(* IEC 61131-3 sources: Elmo_Master/Lasal_PRG/Welcon8Axis_EtherCAT_Test_With_RobotAxis/Network/Robot_Network, 1 file *)

(* ---- ONE_Robot_Network_Table.st ---- *)
#define OBJECTS_CONFIG

//Define part of class _LMCBeltAxis
//#define _DEBUG_MODUS_ISSYNCHRON
//#define _DEBUG_MODUS_CHECKSWLIMIT

#define _LMCBELT_MIN_POS       -16#6FFFFFFF    // default MINPOS when INITvalue=0
#define _LMCBELT_MAX_POS        16#6FFFFFFF    // default MAXPOS when INITvalue=0
#define _LMCBELT_OVERVFLOW_POS  16#7FFFFFFF    // MAX POSITION for checking overflow

#define _LMCBELT_AMAX_SET 2000000000
#define _LMCBELT_VMAX_SET 500000000

//////////////////////
// ruckbegrenzter Modus _JERK_PROFILE
#define LMCBELT_MIN_SHRINK_FACTOR_4_CORRECTTOEXACTPOS 0.9
#define LMCBELT_MAX_SHRINK_FACTOR_4_CORRECTTOEXACTPOS_FAR 1.2
#define LMCBELT_MAX_SHRINK_FACTOR_4_CORRECTTOEXACTPOS_NEAR 5.0
#define LMCBELT_MAX_SHRINK_FACTOR_4_CORRECTTOEXACTPOS_WINDOW 5.0

#define LMCBELT_MAX_TIME_TO_WAIT_4_BRAKING 3.0 //in Ticks
#define LMCBELT_MAX_DURATION_WITH_MAX_ACCEL_TO_MASTER 20000  //in Ticks
#define LMCBELT_ALLOWED_AJMP_FACTOR 1.1
#define LMCBELT_FACTOR_4_ALLOWED_MASTER_ACCEL_PROFILE_COUPLING 1.2
#define LMCBELT_ACCEL_FACTOR_4_PROFILE_COUPLING 1.1
#define LMCBELT_JERK_FACTOR_4_PROFILE_COUPLING 1.2
#define LMCBELT_FACTOR_2_REDUCE_AXIS_ACC_LIMIT 1.02

//////////////////////
// LREAL Modi
// #define DEBUG_TRAP_DELTA_ACCEL
#define _LMCBELT_LREAL_EPSILON 0.000001

#ifndef _DINT_MIN
#define _DINT_MIN -2147483648
#endif

#ifndef _DINT_MAX
#define _DINT_MAX 2147483647
#endif

#define _LMCBELT_MIN_VEL_MOVECMD 1 // minimale programmierbare Geschwindigkeit für LREAL-MoveTypes [internal units / sec]
#include <.\lsl_st_systrace.h>
#include "..\..\Class\_LMCAxisBase\C_MathAxis.h"
#include "..\..\Class\_LMCAxisBase\_LMCTraceView.h"
//Define part of class _LMCMath_SO3
// maximal inaccuracies of LREAL
#define _LREAL_EPSILON        0.000001
#define _LREAL_EPSILON_MUL    0.000001
// minmal volume of orthogonalsystem
#define MIN_SPAT_PRODUCT      _LREAL_EPSILON_MUL

#ifndef deg
  #define SCALE_ROT_ANGLE       (10000)
#else
  #define SCALE_ROT_ANGLE       (1deg)
#endif

#define SCALE_VECTOR          (10000)
//Define part of class _LMCMathFunctions
#define _INT_DEG                       * 1024 * 1000 //Internal Resolution of Degrees
#define LMC_PI                          3.1415926535897932384626433832795   //LMC_ avoids name clash

#define _LMC_EPSILON    0.000001
#define _MATH_EPSILON   0.000000001

//LREAL Zero Test:
#ifndef _LMCMATH_FLOAT_ISZERO
  #define _LMCMATH_FLOAT_ISZERO(p1)            ((p1 > -_LMC_EPSILON) & (p1 < _LMC_EPSILON))
#endif
#ifndef _LMCMATH_FLOAT_NOTZERO
  #define _LMCMATH_FLOAT_NOTZERO(p1)           ((p1 < -_LMC_EPSILON) | (p1 > _LMC_EPSILON))
#endif
#ifndef _LMCMATH_FLOAT_EQUAL
  #define _LMCMATH_FLOAT_EQUAL(p1,p2)          (((p1 - p2) < _LMC_EPSILON) & ((p1 - p2) > -_LMC_EPSILON))
#endif

#define _LMCMATH_LREAL_MAX  1.79E308
#define _LMCMATH_REAL_MAX   3.4E38

#ifndef _DINT_MIN
  #define _DINT_MIN -2147483648
#endif

#define LMC_NUMERIC_TOLERANCE   (0.000000001)
#define LMC_RESOLVE_TOLERANCE       (0.000000001)

// 25µsec für ein repeat auf ARM CP 111
#define LMC_MAX_REPEAT      25

// Geschwindigkeit wird auf 1 interne Einheit genau iteriert
#define PRECIS_REPEAT   (1.0)

//#define INTERN_MATH_TEST
#include "..\..\Class\_LMCMathFunctions\C_MathFunct.h"
//Define part of class _LMCProfileBase
#pragma once

// DEBUG MODUS TO DEACTIVATE ACTIVE MUTEX
//#define DEBUG_MODUS
//#define DEBUG_CMD_TYPE

#pragma once

//LREAL Zero Test:
#ifndef _LMCPROF_LREAL_ISZERO
  #define _LMCPROF_LREAL_ISZERO(p1)           ((p1 > -_LMCPROF_EPSILON) & (p1 < _LMCPROF_EPSILON))
#endif
#ifndef _LMCPROF_LREAL_NOTZERO
  #define _LMCPROF_LREAL_NOTZERO(p1)          ((p1 < -_LMCPROF_EPSILON) | (p1 > _LMCPROF_EPSILON))
#endif
#define _LMCPROF_LREAL_MAX                    1.79E308

#define _LMPROF_PROMILLE                      1000

//Move Curve Spline Defines
#define _LMC_PROF_MCS_MINOVERDRIVE                -900
#define _LMC_PROF_MCS_MAXOVERDRIVE                10000 //=> Centripetal Acceleration can be up to 10 * given AMove
#define _LMC_PROF_MCS_DEFAULT_JERKSMOOTH          1

#define _LMC_PROF_CES_DEFAULT_ZEXPONENT           1.0 //Default Spline Z Exponent used in calcEllipseSpline(), set with SetProfileParameter()
#define _LMC_PROF_CES_MAX_ZEXPONENT_W_LIN         1.0 //Max Spline Z Exponent if moving with Linear movements, used in calcEllipseSpline()
#define _LMC_PROF_CES_MIN_ZEXPONENT               1.0 //Min Spline Z Exponent, used in calcEllipseSpline()

#define _LMC_PROF_ERRORBUFFER_ENTRIES             10
#define _LMC_PROF_MAINGROUP                       1 // Achse ist in Hauptgruppe
#define _LMC_PROF_SLAVEGROUP1                     2 // Achse ist in Nebengruppe 1
#define _LMC_PROF_SLAVEGROUP2                     3 // Achse ist in Nebengruppe 2
#define _LMC_PROF_SLAVEGROUP3                     4 // Achse ist in Nebengruppe 3
#define _LMC_PROF_SLAVEGROUP4                     5 // Achse ist in Nebengruppe 4
#define _LMC_PROF_SLAVEGROUP5                     6 // Achse ist in Nebengruppe 5

#define _LMC_PROF_MAX_SLAVEGROUPS               _LMC_PROF_SLAVEGROUP5

#define _LMCPROF_NEEDED_FREE_BUFFER_ENTRIES    4

#define _LMC_PROF_MAXOVERRIDE	               1000 // Maximalwert für Override
#define _LMC_PROF_MINOVERRIDE	                  0	// Minimalwert für Override
#define _LMC_PROF_NORMOVERRIDE               1000 // 100%-Wert für Override

#define _LMC_PROF_MAX_DINT                   2147483647
#define _LMC_PROF_MAX_UDINT                  4294967295

#define TRANS1                                  0 //index of 1. transition elmt
#define TRANS2                                  1 //index of 2. transition elmt
#define TRANS3                                  2 //index of 3. transition elmt

#define _LMC_PROF_VECTOR_WINDOW                 10mm

#define MIN_TRANSRAD_PPTH                       0
#define DEF_TRANSRAD_PPTH                       500
#define MOVECURVE_ACCEL_PATH_AUXAXIS            250 // 250 // 25% of the path length is used for accelerating auxiliary axes with splines

#define _LMC_PROF_DEFAULT_MAX_TANG_ERR          900000 //90° ist defaultmäßig maximale tangential fehler

#define _LMC_PROF_RESTARTPROF_TOLSPHERE_DEFAULT 1mm
#define _LMC_PROF_RESTARTPROF_APPROACH_DEFAULT  0

#define _LMC_PROF_MULT_LOOKAHEAD_LINE           5 //default multiplier for lookaheadsmalllines

#define _LMCPROF_REDUCEMOVINGTIME_MAXFACTOR  10000

// the minimal height difference between the end / beginning of the linear part of a MoveCurve() movement and the start / end of the MoveCurveAux section
#define _LMCPROF_MINIMAL_SWERVEDIFF            0.2mm

// Fehlertoleranz bei Umrechnung von Integer auf Float
#define RESOLUTION_ERROR      (5.0)
// Fehlertoleranz wenn der Ruck innerhalb eines Ticks um 2*Jmax springt
#define JERKTICK_ERROR        (-1.0)

// Rückgabeparameter
#define CALCRESIDT_NO_ERROR            0
#define CALCRESIDT_INIT_ERROR          -1
#define CALCRESIDT_NO_SOLUTION         -2

// Präfix (wird für Ruck verwendet)
#ifndef PREFIX_KILO
  #define PREFIX_KILO             (1000.0)
#endif
// Umrechnung von Sekunden auf Ticks
#ifndef CONVERT_SEC_TO_MSEC
  #define CONVERT_SEC_TO_MSEC   (1000.0)
#endif
// interne Mathematik-Tests - speziell Genauigkeitstest von LREAL
//#define INTERN_TEST

// =======================================================
// Defines for Clothoid (Parameters / Conversion)
// Minimal angle to use a compound solution
#define _LMCPROF_CLOTH_MINTAU                  0.06        // 0.06 (radiant) = R/3 clothoid identification
#define _LMCPROF_CLOTH_HAIRPINLIMIT            0.0004      // 0.0004 (radiant) < 0.025 degree - Limit, when the turn is close to a hairpin (cone angle smaller than this limit - handle it is a stop)
#define _LMCPROF_CLOTH_TABLESCALE              0.000000001 // 10^(-9) // This value is a fixed scale of the unit cloth table - when this value is changed, the table must be changed too.

//Angle conversion
#ifndef _LMCPROF_DEG_RAD
  #define _LMCPROF_DEG_RAD(p1)       (((p1) / (180.0 * 1deg)) * _PI)
#endif
#ifndef _LMCPROF_RAD_DEG
  #define _LMCPROF_RAD_DEG(p1)       (((p1) / _PI) * 180.0) * 1deg
#endif

// Defines for tangential axis
#define _LMCPROF_TANGAXIS_ACTANGLEOVERFLOWLIMIT    45.0 deg
#define _LMCPROF_TANGAXIS_OVERFLOWDETECTLIMIT     359.0 deg

// Maximum allowed number of points per spline -
// Attention! If this value is changed also the MaxNrOfPointsPerMoveMaxValue of MoveSplineTable and
// IPR_MAX_NR_SPLINE_POINTS of _LMCCNCIPRBase are to be changed
#define PROF_MAX_NR_SPLINE_POINTS           50
// Maximal number of spline points is twice as high as the number of points - 1 (movement to the last point can't include addition intermediate move)
#define PROF_MaxNrSplineTargets             ((PROF_MAX_NR_SPLINE_POINTS * 2) - 1)

// Move Spline minimal trajectory angle
#define _LMC_PROF_MOVESPLINE_MIN_ANGLE      45 deg // 45 deg
#include "..\..\Class\_LMCProfileBase\C_MathProfile.h"
//Define part of class _LMCProfileBuffer
#define    _LMC_PB_MINENTRIES     201
#define    _LMC_PB_MAXENTRIES     2000

#define _LMC_PB_TMP_MINENTRIES    7
#define _LMC_PB_TMP_MAXENTRIES    100

#define _LMC_PB_RB_MINENTRIES     5
#define _LMC_PB_RB_MAXENTRIES     10

//////////////////////
// Mutex
#define MUTEX_NAME_MAX_LENGTH_LMCPROFILE     32   //maximale Anzahl an Zeichen für den Mutexnamen
#define MUTEX_NAME_END_LENGTH_LMCPROFILE      3
#define STR_MUTEX_NAME_SEPERATOR_LMCPROFILE ".."
//Define part of class _LMCRobotBase
#define DELAYPOWERONHWAXES_TIMEOUT        0
#define DELAYPOWEROFF_TIMEOUT             0
#define WAITPOWERONHWAXES_TIMEOUT     30sec
#define CHECKREFERENCEHWAXES_TIMEOUT  30sec
#define WAITPOWERONKINAXES_TIMEOUT    30sec
#define CHECKCOUPLEHWAXES_TIMEOUT        50
#define WAITPROFILESTOPPED_TIMEOUT     1000
#define WAITSTOPMOVEKINAXES_TIMEOUT    1000
#define WAITSTOPMOVEHWAXES_TIMEOUT     1000
#define WAITERRORQUIT_TIMEOUT           800

#define STOPMOVEPOSITIONWINDOW_DEFAULT 1mm
#define START_COUPLEWINDOW_DEFAULT     1mm

#define GET_LINE_OFFSET 1000000

#define ALL_HW_AXES -1
#define ALL_KINEMATIC_AXES -2
#define ALL_PROFILE_AXES -3
#define ALL_AXES_101_TO_109 -4
#define ALL_ROBOT_AXES 0

#define SCALE_ROTAXIS 100000
#define SCALE_KOFAC 1000000

#define LIMIT_BELT_CMD            2
#define SYNC_DESYNC_FULL_LENGTH   1000

#define SYNC_DESYNC_MIN_LENGTH      50

#define BELTCOUPLING_DEFAULT_FILTER_DEPTH_VMASTER 40 //Bei Änderungen auch Kommentar von _LMCROBOT_BELTCOUPLING_VEL_FILTER_DEPTH anpassen!
#define BELTCOUPLING_MAX_FILTER_DEPTH_VMASTER 60 //Bei Änderungen auch Kommentar von _LMCROBOT_BELTCOUPLING_VEL_FILTER_DEPTH anpassen!

#define ROTATORY_DISK_MODULO (360deg)
#define ROTATORY_DISK_ANGLE_TO_RADIANT (2.0*LMC_PI/(ROTATORY_DISK_MODULO))

#ifndef CIRCLE3D_NO_HELIX_MAX_DEVIATION
  #define CIRCLE3D_NO_HELIX_MAX_DEVIATION 0.02
#endif
//Define part of class _LMCSplineBuffer
#define LMCSPLINEBUFF_MINBUFFS              3             //SplineGroups
#define LMCSPLINEBUFF_EPSILON               0.000001
#define LMCSPLINEBUFF_MAX_SPLINES_PER_GROUP 40
#define LMCSPLINEBUFF_MALLOC_MARK           9
#define LMCSPLINEBUFF_HIRES_VEL_DEFAULT     (1000.0)
#define LMCSPLINEBUFF_HIRES_ACC_DEFAULT     (10000.0)
#define LMCSPLINEBUFF_HIRES_JERK_DEFAULT    (1000000.0)
#define LMCSPLINEBUFF_CALCPARAS_POS         16#00000001
#define LMCSPLINEBUFF_CALCPARAS_VEL         16#00000002
#define LMCSPLINEBUFF_CALCPARAS_ACC         16#00000004
#define LMCSPLINEBUFF_CALCPARAS_JERK        16#00000008
#define LMCSPLINEBUFF_CALCPARAS_JOUNCE      16#00000010
#define LMCSPLINEBUFF_SEARCH_ITER_DEFAULT   100
#define LMCSPLINEBUFF_SEARCH_WIN_DEFAULT    1.0

//Coeffecient Short Names:
#define SB_CO_A (pSplineSection^.Coefficients.lrCoefficient1)
#define SB_CO_B (pSplineSection^.Coefficients.lrCoefficient2)
#define SB_CO_C (pSplineSection^.Coefficients.lrCoefficient3)
#define SB_CO_D (pSplineSection^.Coefficients.lrCoefficient4)
#define SB_CO_E (pSplineSection^.Coefficients.lrCoefficient5)
#define SB_CO_F (pSplineSection^.Coefficients.lrCoefficient6)
#define SB_CO_G (pSplineSection^.Coefficients.lrCoefficient7)
#define SB_CO_H (pSplineSection^.Coefficients.lrCoefficient8)
#define SB_TICK (pSplineSection^.lrTick)
//Define part of class _LMCTableBuffer
#define _TABLE_POINT_COUNT_ 100

#define _TABLE_POINT_20PERCENT 25
#define _TABLE_POINT_35PERCENT 40
#define _TABLE_POINT_50PERCENT 50
#define _TABLE_POINT_65PERCENT 60
#define _TABLE_POINT_80PERCENT 75

#define _LMCTABLEBUFFER_MALLOCMARK  9

FUNCTION GLOBAL TAB ONE_Robot_Network
-1$UINT, 0$UINT,
0$UINT, 0$UINT,

16$UDINT,
TO_UDINT(1064285160), "_LMCBeltAxis", 1$UINT, 7$UINT, 1$UINT,
TO_UDINT(4293818033), "_LMCMath_SO3", 1$UINT, 24$UINT, 2$UINT,
TO_UDINT(838927485), "_LMCMathFunctions", 1$UINT, 75$UINT, 2$UINT,
TO_UDINT(2952189205), "_LMCProfile", 3$UINT, 0$UINT, 0$UINT,
TO_UDINT(506182625), "_LMCProfileBase", 4$UINT, 0$UINT, 0$UINT,
TO_UDINT(2726627155), "_LMCProfileBuffer", 1$UINT, 53$UINT, 1$UINT,
TO_UDINT(2883857672), "_LMCProfileLog", 1$UINT, 44$UINT, 1$UINT,
TO_UDINT(4141185109), "_LMCProfileVis", 1$UINT, 30$UINT, 1$UINT,
TO_UDINT(3174746949), "_LMCProfileVisAxis", 1$UINT, 20$UINT, 9$UINT,
TO_UDINT(4192117043), "_LMCProfileVisInt", 1$UINT, 41$UINT, 1$UINT,
TO_UDINT(1543035932), "_LMCProfileVisMovePara", 1$UINT, 30$UINT, 6$UINT,
TO_UDINT(3888346726), "_LMCRobotBase", 2$UINT, 22$UINT, 1$UINT,
TO_UDINT(4210476436), "_LMCRobotLog", 1$UINT, 42$UINT, 1$UINT,
TO_UDINT(1286231841), "_LMCSplineBuffer", 1$UINT, 2$UINT, 1$UINT,
TO_UDINT(2328372307), "_LMCTableBuffer", 1$UINT, 23$UINT, 1$UINT,
TO_UDINT(1472648579), "Robot_Handler", 0$UINT, 0$UINT, 1$UINT,

1$UINT, TO_UDINT(3188917884), "_LMCROBOTBASE1\LMCBELTINTERNAL",

1$UINT, TO_UDINT(2922016232), "_LMCROBOTBASE1\LMCMATH_SO3",
1$UINT, TO_UDINT(1366148008), "_LMCROBOTBASE1\_BASE\_LMCMATH_SO3",

1$UINT, TO_UDINT(1157192838), "_LMCROBOTBASE1\LMCBELTINTERNAL\LMCMATH",
1$UINT, TO_UDINT(2796190616), "_LMCROBOTBASE1\_BASE\_LMCMATHFUNCTIONS",

1$UINT, TO_UDINT(909015222), "_LMCROBOTBASE1\_BASE\_LMCPROFILEBUFFER",

1$UINT, TO_UDINT(2347724176), "_LMCROBOTBASE1\_BASE\_LMCPROFILELOG",

1$UINT, TO_UDINT(3604887757), "_LMCROBOTBASE1\_BASE\_LMCPROFILEVIS",

1$UINT, TO_UDINT(4143639116), "_LMCROBOTBASE1\_BASE\_LMCPROFILEVIS\_LMCPROFILEVISAXIS1",
1$UINT, TO_UDINT(1878244342), "_LMCROBOTBASE1\_BASE\_LMCPROFILEVIS\_LMCPROFILEVISAXIS2",
1$UINT, TO_UDINT(418679648), "_LMCROBOTBASE1\_BASE\_LMCPROFILEVIS\_LMCPROFILEVISAXIS3",
1$UINT, TO_UDINT(2257592003), "_LMCROBOTBASE1\_BASE\_LMCPROFILEVIS\_LMCPROFILEVISAXIS4",
1$UINT, TO_UDINT(4053216853), "_LMCROBOTBASE1\_BASE\_LMCPROFILEVIS\_LMCPROFILEVISAXIS5",
1$UINT, TO_UDINT(1755217903), "_LMCROBOTBASE1\_BASE\_LMCPROFILEVIS\_LMCPROFILEVISAXIS6",
1$UINT, TO_UDINT(530141049), "_LMCROBOTBASE1\_BASE\_LMCPROFILEVIS\_LMCPROFILEVISAXIS7",
1$UINT, TO_UDINT(2401653480), "_LMCROBOTBASE1\_BASE\_LMCPROFILEVIS\_LMCPROFILEVISAXIS8",
1$UINT, TO_UDINT(4162937470), "_LMCROBOTBASE1\_BASE\_LMCPROFILEVIS\_LMCPROFILEVISAXIS9",

1$UINT, TO_UDINT(2979030242), "_LMCROBOTBASE1\_BASE\_LMCPROFILEVIS\_LMCPROFILEVISINT",

1$UINT, TO_UDINT(1783828595), "_LMCROBOTBASE1\_BASE\_LMCPROFILEVIS\_LMCPROFILEVISMOVEPARA1",
1$UINT, TO_UDINT(4082778569), "_LMCROBOTBASE1\_BASE\_LMCPROFILEVIS\_LMCPROFILEVISMOVEPARA2",
1$UINT, TO_UDINT(2220716383), "_LMCROBOTBASE1\_BASE\_LMCPROFILEVIS\_LMCPROFILEVISMOVEPARA3",
1$UINT, TO_UDINT(440001788), "_LMCROBOTBASE1\_BASE\_LMCPROFILEVIS\_LMCPROFILEVISMOVEPARA4",
1$UINT, TO_UDINT(1832834154), "_LMCROBOTBASE1\_BASE\_LMCPROFILEVIS\_LMCPROFILEVISMOVEPARA5",
1$UINT, TO_UDINT(4097279440), "_LMCROBOTBASE1\_BASE\_LMCPROFILEVIS\_LMCPROFILEVISMOVEPARA6",

_NO_ATTR, TO_UDINT(669706412), "_LMCROBOTBASE1",

1$UINT, TO_UDINT(2991295094), "_LMCROBOTBASE1\_LMCROBOTLOG",

1$UINT, TO_UDINT(2213426856), "_LMCROBOTBASE1\_BASE\_LMCSPLINEBUFFER",

1$UINT, TO_UDINT(1950102629), "_LMCROBOTBASE1\_BASE\_LMCTABLEBUFFER",

_NO_ATTR, TO_UDINT(4147837944), "ROBOT_HANDLER1",

//Internal connections
0$UDINT,
27$UDINT,
TO_UDINT(0), "LMCMath", TO_UDINT(3),
TO_UDINT(7), "_LMCProfileVisMovePara1", TO_UDINT(18),
TO_UDINT(7), "_LMCProfileVisMovePara2", TO_UDINT(19),
TO_UDINT(7), "_LMCProfileVisMovePara3", TO_UDINT(20),
TO_UDINT(7), "_LMCProfileVisMovePara4", TO_UDINT(21),
TO_UDINT(7), "_LMCProfileVisMovePara5", TO_UDINT(22),
TO_UDINT(7), "_LMCProfileVisMovePara6", TO_UDINT(23),
TO_UDINT(7), "_LMCProfileVisAxis1", TO_UDINT(8),
TO_UDINT(7), "_LMCProfileVisAxis2", TO_UDINT(9),
TO_UDINT(7), "_LMCProfileVisAxis3", TO_UDINT(10),
TO_UDINT(7), "_LMCProfileVisAxis4", TO_UDINT(11),
TO_UDINT(7), "_LMCProfileVisAxis5", TO_UDINT(12),
TO_UDINT(7), "_LMCProfileVisAxis6", TO_UDINT(13),
TO_UDINT(7), "_LMCProfileVisInt", TO_UDINT(17),
TO_UDINT(7), "_LMCProfileVisAxis7", TO_UDINT(14),
TO_UDINT(7), "_LMCProfileVisAxis8", TO_UDINT(15),
TO_UDINT(7), "_LMCProfileVisAxis9", TO_UDINT(16),
TO_UDINT(24), "_LMCMathFunctions", TO_UDINT(4),
TO_UDINT(24), "_LMCProfileBuffer", TO_UDINT(5),
TO_UDINT(24), "_LMCProfileVis", TO_UDINT(7),
TO_UDINT(24), "_LMCProfileLog", TO_UDINT(6),
TO_UDINT(24), "_LMCTableBuffer", TO_UDINT(27),
TO_UDINT(24), "_LMCSplineBuffer", TO_UDINT(26),
TO_UDINT(24), "_LMCMath_SO3", TO_UDINT(2),
TO_UDINT(24), "LMCMath_SO3", TO_UDINT(1),
TO_UDINT(24), "_LMCRobotLog", TO_UDINT(25),
TO_UDINT(24), "LMCBeltInternal", TO_UDINT(0),
0$UDINT,
23$UDINT,
TO_UDINT(7), "coLMCProfileBase", TO_UDINT(24), "Control",
TO_UDINT(17), "coLMCProfileVisAxis1", TO_UDINT(8), "AxisConnected",
TO_UDINT(17), "coLMCProfileVisAxis2", TO_UDINT(9), "AxisConnected",
TO_UDINT(17), "coLMCProfileVisAxis3", TO_UDINT(10), "AxisConnected",
TO_UDINT(17), "coLMCProfileVisAxis4", TO_UDINT(11), "AxisConnected",
TO_UDINT(17), "coLMCProfileVisAxis5", TO_UDINT(12), "AxisConnected",
TO_UDINT(17), "coLMCProfileVisAxis6", TO_UDINT(13), "AxisConnected",
TO_UDINT(17), "coLMCProfileVisAxis7", TO_UDINT(14), "AxisConnected",
TO_UDINT(17), "coLMCProfileVisAxis8", TO_UDINT(15), "AxisConnected",
TO_UDINT(17), "coLMCProfileVisAxis9", TO_UDINT(16), "AxisConnected",
TO_UDINT(17), "LMCProfileVisMovePara1", TO_UDINT(18), "ClassSvr",
TO_UDINT(17), "LMCProfileVisMovePara2", TO_UDINT(19), "ClassSvr",
TO_UDINT(17), "LMCProfileVisMovePara3", TO_UDINT(20), "ClassSvr",
TO_UDINT(17), "LMCProfileVisMovePara4", TO_UDINT(21), "ClassSvr",
TO_UDINT(17), "LMCProfileVisMovePara5", TO_UDINT(22), "ClassSvr",
TO_UDINT(17), "LMCProfileVisMovePara6", TO_UDINT(23), "ClassSvr",
TO_UDINT(24), "LMCMathFunction", TO_UDINT(4), "ClassSvr",
TO_UDINT(24), "LMCProfileBuffer", TO_UDINT(5), "ClassSvr",
TO_UDINT(24), "LMCLog", TO_UDINT(6), "ClassSvr",
TO_UDINT(24), "LMCTableBuffer", TO_UDINT(27), "TableSize",
TO_UDINT(24), "LMCSplineBuffer", TO_UDINT(26), "ClassSvr",
TO_UDINT(24), "LMCMathSO3", TO_UDINT(2), "Control",
TO_UDINT(28), "RobotBase", TO_UDINT(24), "Control",

//Initialization values
0$UDINT,
32$UDINT,
TO_UDINT(0), "SWMinPos", TO_UDINT(0),//|Robot_Network._LMCRobotBase1\LMCBeltInternal.SWMinPos;
TO_UDINT(0), "SWMaxPos", TO_UDINT(0),//|Robot_Network._LMCRobotBase1\LMCBeltInternal.SWMaxPos;
TO_UDINT(8), "AxisGroup", TO_UDINT(1),//|Robot_Network._LMCProfileVis\_base\_LMCRobotBase1\_LMCProfileVisAxis1.AxisGroup;
TO_UDINT(9), "AxisGroup", TO_UDINT(1),//|Robot_Network._LMCProfileVis\_base\_LMCRobotBase1\_LMCProfileVisAxis2.AxisGroup;
TO_UDINT(10), "AxisGroup", TO_UDINT(1),//|Robot_Network._LMCProfileVis\_base\_LMCRobotBase1\_LMCProfileVisAxis3.AxisGroup;
TO_UDINT(11), "AxisGroup", TO_UDINT(1),//|Robot_Network._LMCProfileVis\_base\_LMCRobotBase1\_LMCProfileVisAxis4.AxisGroup;
TO_UDINT(12), "AxisGroup", TO_UDINT(1),//|Robot_Network._LMCProfileVis\_base\_LMCRobotBase1\_LMCProfileVisAxis5.AxisGroup;
TO_UDINT(13), "AxisGroup", TO_UDINT(1),//|Robot_Network._LMCProfileVis\_base\_LMCRobotBase1\_LMCProfileVisAxis6.AxisGroup;
TO_UDINT(14), "AxisGroup", TO_UDINT(1),//|Robot_Network._LMCProfileVis\_base\_LMCRobotBase1\_LMCProfileVisAxis7.AxisGroup;
TO_UDINT(15), "AxisGroup", TO_UDINT(1),//|Robot_Network._LMCProfileVis\_base\_LMCRobotBase1\_LMCProfileVisAxis8.AxisGroup;
TO_UDINT(16), "AxisGroup", TO_UDINT(1),//|Robot_Network._LMCProfileVis\_base\_LMCRobotBase1\_LMCProfileVisAxis9.AxisGroup;
TO_UDINT(24), "OpMode", TO_UDINT(_LMC_AUTOMATIC),//|Robot_Network._LMCRobotBase1.OpMode;
TO_UDINT(24), "Resolution", TO_UDINT(1),//|Robot_Network._LMCRobotBase1.Resolution;
TO_UDINT(24), "MoveType", TO_UDINT(RAMP_PROFILE),//|Robot_Network._LMCRobotBase1.MoveType;
TO_UDINT(24), "ErrorConfig", TO_UDINT(2#0000000),//|Robot_Network._LMCRobotBase1.ErrorConfig;
TO_UDINT(24), "SimulateMode", TO_UDINT(0),//|Robot_Network._LMCRobotBase1.SimulateMode;
TO_UDINT(24), "VMax", TO_UDINT(5000 mm),//|Robot_Network._LMCRobotBase1.VMax;
TO_UDINT(24), "AMax", TO_UDINT(5000 mm),//|Robot_Network._LMCRobotBase1.AMax;
TO_UDINT(24), "JMax", TO_UDINT(5000 mm),//|Robot_Network._LMCRobotBase1.JMax;
TO_UDINT(26), "No", TO_UDINT(LMCSPLINEBUFF_MINBUFFS),//|Robot_Network._base\_LMCRobotBase1\_LMCSplineBuffer.No;
TO_UDINT(27), "No", TO_UDINT(2),//|Robot_Network._base\_LMCRobotBase1\_LMCTableBuffer.No;
TO_UDINT(28), "Pos1", TO_UDINT(100 mm),//|Robot_Network.Robot_Handler1.Pos1;
TO_UDINT(28), "Pos2", TO_UDINT(100 mm),//|Robot_Network.Robot_Handler1.Pos2;
TO_UDINT(28), "Pos3", TO_UDINT(100 mm),//|Robot_Network.Robot_Handler1.Pos3;
TO_UDINT(28), "Pos4", TO_UDINT(100 mm),//|Robot_Network.Robot_Handler1.Pos4;
TO_UDINT(28), "Pos5", TO_UDINT(100 mm),//|Robot_Network.Robot_Handler1.Pos5;
TO_UDINT(28), "Pos6", TO_UDINT(100 mm),//|Robot_Network.Robot_Handler1.Pos6;
TO_UDINT(28), "Pos7", TO_UDINT(100 mm),//|Robot_Network.Robot_Handler1.Pos7;
TO_UDINT(28), "Pos8", TO_UDINT(100 mm),//|Robot_Network.Robot_Handler1.Pos8;
TO_UDINT(28), "Velo", TO_UDINT(10 mm),//|Robot_Network.Robot_Handler1.Velo;
TO_UDINT(28), "Acc", TO_UDINT(10 mm),//|Robot_Network.Robot_Handler1.Acc;
TO_UDINT(28), "Jerk", TO_UDINT(10 mm),//|Robot_Network.Robot_Handler1.Jerk;

//Symbolic initialization values
0$UDINT,
0$UDINT,

//Initialization of string values
0$UDINT,
0$UDINT,

//Configuration of tasks (RealTime, Cyclic, Background)
0$UDINT,
1$UDINT,
TO_UDINT(24), (1)$UDINT, 4194303$DINT, 	//_LMCROBOTBASE1

0$UDINT,
1$UDINT,
TO_UDINT(24), (1)$UDINT, 4194303$DINT, 	//_LMCROBOTBASE1

0$UDINT,
1$UDINT,
TO_UDINT(17), (500)$UDINT, 4194303$DINT, 	//_LMCROBOTBASE1\_BASE\_LMCPROFILEVIS\_LMCPROFILEVISINT

//External connections
0$UDINT,
8$UDINT,
TO_UDINT(24), "LMCAxis1", C_TRY, TO_UDINT(3550025316), "_LMCAxis_Axis1","Control",
TO_UDINT(24), "LMCAxis2", C_TRY, TO_UDINT(1250969566), "_LMCAxis_Axis2","Control",
TO_UDINT(24), "LMCAxis3", C_TRY, TO_UDINT(1033336648), "_LMCAxis_Axis3","Control",
TO_UDINT(24), "LMCAxis4", C_TRY, TO_UDINT(2750669547), "_LMCAxis_Axis4","Control",
TO_UDINT(24), "LMCAxis5", C_TRY, TO_UDINT(3572814461), "_LMCAxis_Axis5","Control",
TO_UDINT(24), "LMCAxis6", C_TRY, TO_UDINT(1308459975), "_LMCAxis_Axis6","Control",
TO_UDINT(24), "LMCAxis7", C_TRY, TO_UDINT(989508433), "_LMCAxis_Axis7","Control",
TO_UDINT(24), "LMCAxis8", C_TRY, TO_UDINT(2856693440), "_LMCAxis_Axis8","Control",

//Magic internal connections
0$UDINT,
73$UDINT,
TO_UDINT(7), "coLMCAxis1", TO_UDINT(24), "LMCAxis1",
TO_UDINT(7), "coLMCAxis2", TO_UDINT(24), "LMCAxis2",
TO_UDINT(7), "coLMCAxis3", TO_UDINT(24), "LMCAxis3",
TO_UDINT(7), "coLMCAxis4", TO_UDINT(24), "LMCAxis4",
TO_UDINT(7), "coLMCAxis5", TO_UDINT(24), "LMCAxis5",
TO_UDINT(7), "coLMCAxis6", TO_UDINT(24), "LMCAxis6",
TO_UDINT(7), "coLMCAxis7", TO_UDINT(24), "LMCAxis7",
TO_UDINT(7), "coLMCAxis8", TO_UDINT(24), "LMCAxis8",
TO_UDINT(7), "coLMCAxis9", TO_UDINT(24), "LMCAxis9",
TO_UDINT(8), "coLMCAxis", TO_UDINT(7), "coLMCAxis1",
TO_UDINT(9), "coLMCAxis", TO_UDINT(7), "coLMCAxis2",
TO_UDINT(10), "coLMCAxis", TO_UDINT(7), "coLMCAxis3",
TO_UDINT(11), "coLMCAxis", TO_UDINT(7), "coLMCAxis4",
TO_UDINT(12), "coLMCAxis", TO_UDINT(7), "coLMCAxis5",
TO_UDINT(13), "coLMCAxis", TO_UDINT(7), "coLMCAxis6",
TO_UDINT(14), "coLMCAxis", TO_UDINT(7), "coLMCAxis7",
TO_UDINT(15), "coLMCAxis", TO_UDINT(7), "coLMCAxis8",
TO_UDINT(16), "coLMCAxis", TO_UDINT(7), "coLMCAxis9",
TO_UDINT(17), "LMCProfileBase", TO_UDINT(7), "coLMCProfileBase",
TO_UDINT(18), "coLMCAxis1", TO_UDINT(7), "coLMCAxis1",
TO_UDINT(18), "coLMCAxis2", TO_UDINT(7), "coLMCAxis2",
TO_UDINT(18), "coLMCAxis3", TO_UDINT(7), "coLMCAxis3",
TO_UDINT(18), "coLMCAxis4", TO_UDINT(7), "coLMCAxis4",
TO_UDINT(18), "coLMCAxis5", TO_UDINT(7), "coLMCAxis5",
TO_UDINT(18), "coLMCAxis6", TO_UDINT(7), "coLMCAxis6",
TO_UDINT(18), "coLMCAxis7", TO_UDINT(7), "coLMCAxis7",
TO_UDINT(18), "coLMCAxis8", TO_UDINT(7), "coLMCAxis8",
TO_UDINT(18), "coLMCAxis9", TO_UDINT(7), "coLMCAxis9",
TO_UDINT(19), "coLMCAxis1", TO_UDINT(7), "coLMCAxis1",
TO_UDINT(19), "coLMCAxis2", TO_UDINT(7), "coLMCAxis2",
TO_UDINT(19), "coLMCAxis3", TO_UDINT(7), "coLMCAxis3",
TO_UDINT(19), "coLMCAxis4", TO_UDINT(7), "coLMCAxis4",
TO_UDINT(19), "coLMCAxis5", TO_UDINT(7), "coLMCAxis5",
TO_UDINT(19), "coLMCAxis6", TO_UDINT(7), "coLMCAxis6",
TO_UDINT(19), "coLMCAxis7", TO_UDINT(7), "coLMCAxis7",
TO_UDINT(19), "coLMCAxis8", TO_UDINT(7), "coLMCAxis8",
TO_UDINT(19), "coLMCAxis9", TO_UDINT(7), "coLMCAxis9",
TO_UDINT(20), "coLMCAxis1", TO_UDINT(7), "coLMCAxis1",
TO_UDINT(20), "coLMCAxis2", TO_UDINT(7), "coLMCAxis2",
TO_UDINT(20), "coLMCAxis3", TO_UDINT(7), "coLMCAxis3",
TO_UDINT(20), "coLMCAxis4", TO_UDINT(7), "coLMCAxis4",
TO_UDINT(20), "coLMCAxis5", TO_UDINT(7), "coLMCAxis5",
TO_UDINT(20), "coLMCAxis6", TO_UDINT(7), "coLMCAxis6",
TO_UDINT(20), "coLMCAxis7", TO_UDINT(7), "coLMCAxis7",
TO_UDINT(20), "coLMCAxis8", TO_UDINT(7), "coLMCAxis8",
TO_UDINT(20), "coLMCAxis9", TO_UDINT(7), "coLMCAxis9",
TO_UDINT(21), "coLMCAxis1", TO_UDINT(7), "coLMCAxis1",
TO_UDINT(21), "coLMCAxis2", TO_UDINT(7), "coLMCAxis2",
TO_UDINT(21), "coLMCAxis3", TO_UDINT(7), "coLMCAxis3",
TO_UDINT(21), "coLMCAxis4", TO_UDINT(7), "coLMCAxis4",
TO_UDINT(21), "coLMCAxis5", TO_UDINT(7), "coLMCAxis5",
TO_UDINT(21), "coLMCAxis6", TO_UDINT(7), "coLMCAxis6",
TO_UDINT(21), "coLMCAxis7", TO_UDINT(7), "coLMCAxis7",
TO_UDINT(21), "coLMCAxis8", TO_UDINT(7), "coLMCAxis8",
TO_UDINT(21), "coLMCAxis9", TO_UDINT(7), "coLMCAxis9",
TO_UDINT(22), "coLMCAxis1", TO_UDINT(7), "coLMCAxis1",
TO_UDINT(22), "coLMCAxis2", TO_UDINT(7), "coLMCAxis2",
TO_UDINT(22), "coLMCAxis3", TO_UDINT(7), "coLMCAxis3",
TO_UDINT(22), "coLMCAxis4", TO_UDINT(7), "coLMCAxis4",
TO_UDINT(22), "coLMCAxis5", TO_UDINT(7), "coLMCAxis5",
TO_UDINT(22), "coLMCAxis6", TO_UDINT(7), "coLMCAxis6",
TO_UDINT(22), "coLMCAxis7", TO_UDINT(7), "coLMCAxis7",
TO_UDINT(22), "coLMCAxis8", TO_UDINT(7), "coLMCAxis8",
TO_UDINT(22), "coLMCAxis9", TO_UDINT(7), "coLMCAxis9",
TO_UDINT(23), "coLMCAxis1", TO_UDINT(7), "coLMCAxis1",
TO_UDINT(23), "coLMCAxis2", TO_UDINT(7), "coLMCAxis2",
TO_UDINT(23), "coLMCAxis3", TO_UDINT(7), "coLMCAxis3",
TO_UDINT(23), "coLMCAxis4", TO_UDINT(7), "coLMCAxis4",
TO_UDINT(23), "coLMCAxis5", TO_UDINT(7), "coLMCAxis5",
TO_UDINT(23), "coLMCAxis6", TO_UDINT(7), "coLMCAxis6",
TO_UDINT(23), "coLMCAxis7", TO_UDINT(7), "coLMCAxis7",
TO_UDINT(23), "coLMCAxis8", TO_UDINT(7), "coLMCAxis8",
TO_UDINT(23), "coLMCAxis9", TO_UDINT(7), "coLMCAxis9",

//Configuration of timeslots of tasks (RealTime, Cyclic)
#ifdef __LSLLDR_TIMESLOTS__
0$UDINT,
0$UDINT,

0$UDINT,
0$UDINT,

#endif //__LSLLDR_TIMESLOTS__

//MultiMaster connections
#ifdef __LSLLDR_MULTIMASTER__
0$UDINT,
0$UDINT,
#endif //__LSLLDR_MULTIMASTER__

//Configuration for task ID (RealTime, CyclicTime)
#ifdef __LSLLDR_TASKID__
"\\\\TASKS2  "
0$UDINT,
1$UDINT,
(0)$UDINT, 	//_LMCROBOTBASE1

0$UDINT,
1$UDINT,
(0)$UDINT, 	//_LMCROBOTBASE1

0$UDINT,
1$UDINT,
(0)$UDINT, 	//_LMCROBOTBASE1\_BASE\_LMCPROFILEVIS\_LMCPROFILEVISINT

#endif //__LSLLDR_TASKID__

END_FUNCTION
